Fanuc KAREL source: kd00028.KL

-- PROVISIONAL review KL for V1013-1; original PC SHA256 bfde906d8939e143df9344bf2a737d3a77658468fcaf4c93969d10176310ff2e
-- Incomplete behavior may be omitted. Consult companion uncertainty JSON. Do not deploy.
PROGRAM KD00028
%NOLOCKGROUP
VAR
  I : INTEGER
  J : INTEGER
  B : BOOLEAN
  R : REAL
  S : STRING[80]
BEGIN
  -- UNRESOLVED_PC offsets 5-21; opcodes 9D,81,18,9D,12,22,9D,13,04
  -- UNRESOLVED_PC offsets 26-30; opcodes 7F
END KD00028
